// TIA Portal V17 export
FUNCTION_BLOCK "FB_T03_Fronts"   // FB103, LAD
{ S7_Optimized_Access := 'TRUE' }
// stored: IsIECCheckEnabled false, MemoryReserve 100, SetENOAutomatically false
   VAR_INPUT
      Capteur : Bool;
   END_VAR
   VAR_OUTPUT
      Impulsion_P : Bool;
      Impulsion_N : Bool;
   END_VAR
   VAR
      Mem_FrontP : Bool;
      Mem_FrontN : Bool;
   END_VAR
   VAR_TEMP   // added for the SCL form of the ladder/FBD networks
      _w1 : Bool;
   END_VAR
BEGIN

REGION Network 1: Front montant
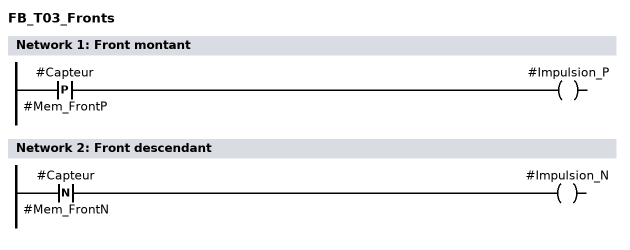
   #_w1 := #Capteur AND NOT #Mem_FrontP;   // rising edge of #Capteur
   #Mem_FrontP := #Capteur;
   #Impulsion_P := #_w1;
END_REGION

REGION Network 2: Front descendant
   #_w1 := NOT #Capteur AND #Mem_FrontN;   // falling edge of #Capteur
   #Mem_FrontN := #Capteur;
   #Impulsion_N := #_w1;
END_REGION
END_FUNCTION_BLOCK
